(* IEC 61131-3 sources: Gen-AI/release/member2-v1.1/成员2_提交包_v1.1/validation/toolchain_smoke_v1.1/C01_undeclared/tools/check/authoritative, 1 file *)

(* ---- source.st ---- *)
FUNCTION_BLOCK FB_AgentProbeUndeclared
VAR_OUTPUT
 y : BOOL;
END_VAR
y := AgentSignalNotDeclared_6E79B1;
END_FUNCTION_BLOCK
